(* IEC 61131-3 sources: llm-plc-st-eval/codesys/dobles/I8, 8 files *)

(* ---- 01_Correcta.st ---- *)
(* DOBLE DE PRUEBA I8/Correcta - NO ES CORPUS. Esperado: veredicto 1 *)
FUNCTION_BLOCK FB_Compresor
VAR_INPUT
    pOilOk : BOOL;
    tempOk : BOOL;
    sinAlm : BOOL;
    btnMarcha : BOOL;
    btnParo : BOOL;
END_VAR
VAR_OUTPUT
    comp : BOOL;
    causaBloqueo : INT;
END_VAR
VAR
    tOil : TON;
    fMarcha : R_TRIG;
    oil : BOOL;
    perm : BOOL;
    lat : BOOL;
    pet : BOOL;
END_VAR
tOil(IN := pOilOk, PT := T#3S);
oil := tOil.Q;
IF NOT oil THEN
    causaBloqueo := 1;
ELSIF NOT tempOk THEN
    causaBloqueo := 2;
ELSIF NOT sinAlm THEN
    causaBloqueo := 3;
ELSE
    causaBloqueo := 0;
END_IF
perm := causaBloqueo = 0;
fMarcha(CLK := btnMarcha);
IF btnParo OR NOT perm THEN
    comp := FALSE;
ELSIF fMarcha.Q THEN
    comp := TRUE;
END_IF
END_FUNCTION_BLOCK

(* ---- 02_SinTemporizacionAceite.st ---- *)
(* DOBLE DE PRUEBA I8/SinTemporizacionAceite - NO ES CORPUS. Esperado: veredicto 2, falla en el paso 1 *)
FUNCTION_BLOCK FB_Compresor
VAR_INPUT
    pOilOk : BOOL;
    tempOk : BOOL;
    sinAlm : BOOL;
    btnMarcha : BOOL;
    btnParo : BOOL;
END_VAR
VAR_OUTPUT
    comp : BOOL;
    causaBloqueo : INT;
END_VAR
VAR
    tOil : TON;
    fMarcha : R_TRIG;
    oil : BOOL;
    perm : BOOL;
    lat : BOOL;
    pet : BOOL;
END_VAR
oil := pOilOk;
IF NOT oil THEN
    causaBloqueo := 1;
ELSIF NOT tempOk THEN
    causaBloqueo := 2;
ELSIF NOT sinAlm THEN
    causaBloqueo := 3;
ELSE
    causaBloqueo := 0;
END_IF
perm := causaBloqueo = 0;
fMarcha(CLK := btnMarcha);
IF btnParo OR NOT perm THEN
    comp := FALSE;
ELSIF fMarcha.Q THEN
    comp := TRUE;
END_IF
END_FUNCTION_BLOCK

(* ---- 03_RearranqueAutomatico.st ---- *)
(* DOBLE DE PRUEBA I8/RearranqueAutomatico - NO ES CORPUS. Esperado: veredicto 2, falla en el paso 6 *)
FUNCTION_BLOCK FB_Compresor
VAR_INPUT
    pOilOk : BOOL;
    tempOk : BOOL;
    sinAlm : BOOL;
    btnMarcha : BOOL;
    btnParo : BOOL;
END_VAR
VAR_OUTPUT
    comp : BOOL;
    causaBloqueo : INT;
END_VAR
VAR
    tOil : TON;
    fMarcha : R_TRIG;
    oil : BOOL;
    perm : BOOL;
    lat : BOOL;
    pet : BOOL;
END_VAR
tOil(IN := pOilOk, PT := T#3S);
oil := tOil.Q;
IF NOT oil THEN
    causaBloqueo := 1;
ELSIF NOT tempOk THEN
    causaBloqueo := 2;
ELSIF NOT sinAlm THEN
    causaBloqueo := 3;
ELSE
    causaBloqueo := 0;
END_IF
perm := causaBloqueo = 0;
fMarcha(CLK := btnMarcha);
lat := (lat OR fMarcha.Q) AND NOT btnParo;
comp := lat AND perm;
END_FUNCTION_BLOCK

(* ---- 04_MarchaPrioritaria.st ---- *)
(* DOBLE DE PRUEBA I8/MarchaPrioritaria - NO ES CORPUS. Esperado: veredicto 2, falla en el paso 7 *)
FUNCTION_BLOCK FB_Compresor
VAR_INPUT
    pOilOk : BOOL;
    tempOk : BOOL;
    sinAlm : BOOL;
    btnMarcha : BOOL;
    btnParo : BOOL;
END_VAR
VAR_OUTPUT
    comp : BOOL;
    causaBloqueo : INT;
END_VAR
VAR
    tOil : TON;
    fMarcha : R_TRIG;
    oil : BOOL;
    perm : BOOL;
    lat : BOOL;
    pet : BOOL;
END_VAR
tOil(IN := pOilOk, PT := T#3S);
oil := tOil.Q;
IF NOT oil THEN
    causaBloqueo := 1;
ELSIF NOT tempOk THEN
    causaBloqueo := 2;
ELSIF NOT sinAlm THEN
    causaBloqueo := 3;
ELSE
    causaBloqueo := 0;
END_IF
perm := causaBloqueo = 0;
fMarcha(CLK := btnMarcha);
IF fMarcha.Q AND perm THEN
    comp := TRUE;
ELSIF btnParo OR NOT perm THEN
    comp := FALSE;
END_IF
END_FUNCTION_BLOCK

(* ---- 05_ArrancaPorNivel.st ---- *)
(* DOBLE DE PRUEBA I8/ArrancaPorNivel - NO ES CORPUS. Esperado: veredicto 2, falla en el paso 8 *)
FUNCTION_BLOCK FB_Compresor
VAR_INPUT
    pOilOk : BOOL;
    tempOk : BOOL;
    sinAlm : BOOL;
    btnMarcha : BOOL;
    btnParo : BOOL;
END_VAR
VAR_OUTPUT
    comp : BOOL;
    causaBloqueo : INT;
END_VAR
VAR
    tOil : TON;
    fMarcha : R_TRIG;
    oil : BOOL;
    perm : BOOL;
    lat : BOOL;
    pet : BOOL;
END_VAR
tOil(IN := pOilOk, PT := T#3S);
oil := tOil.Q;
IF NOT oil THEN
    causaBloqueo := 1;
ELSIF NOT tempOk THEN
    causaBloqueo := 2;
ELSIF NOT sinAlm THEN
    causaBloqueo := 3;
ELSE
    causaBloqueo := 0;
END_IF
perm := causaBloqueo = 0;
fMarcha(CLK := btnMarcha);
comp := (comp OR btnMarcha) AND perm AND NOT btnParo;
END_FUNCTION_BLOCK

(* ---- 06_CausaPrioridadInvertida.st ---- *)
(* DOBLE DE PRUEBA I8/CausaPrioridadInvertida - NO ES CORPUS. Esperado: veredicto 2, falla en el paso 0 *)
FUNCTION_BLOCK FB_Compresor
VAR_INPUT
    pOilOk : BOOL;
    tempOk : BOOL;
    sinAlm : BOOL;
    btnMarcha : BOOL;
    btnParo : BOOL;
END_VAR
VAR_OUTPUT
    comp : BOOL;
    causaBloqueo : INT;
END_VAR
VAR
    tOil : TON;
    fMarcha : R_TRIG;
    oil : BOOL;
    perm : BOOL;
    lat : BOOL;
    pet : BOOL;
END_VAR
tOil(IN := pOilOk, PT := T#3S);
oil := tOil.Q;
IF NOT sinAlm THEN
    causaBloqueo := 3;
ELSIF NOT tempOk THEN
    causaBloqueo := 2;
ELSIF NOT oil THEN
    causaBloqueo := 1;
ELSE
    causaBloqueo := 0;
END_IF
perm := causaBloqueo = 0;
fMarcha(CLK := btnMarcha);
IF btnParo OR NOT perm THEN
    comp := FALSE;
ELSIF fMarcha.Q THEN
    comp := TRUE;
END_IF
END_FUNCTION_BLOCK

(* ---- 07_AceiteNoContinuo.st ---- *)
(* DOBLE DE PRUEBA I8/AceiteNoContinuo - NO ES CORPUS. Esperado: veredicto 2, falla en el paso 12 *)
FUNCTION_BLOCK FB_Compresor
VAR_INPUT
    pOilOk : BOOL;
    tempOk : BOOL;
    sinAlm : BOOL;
    btnMarcha : BOOL;
    btnParo : BOOL;
END_VAR
VAR_OUTPUT
    comp : BOOL;
    causaBloqueo : INT;
END_VAR
VAR
    tOil : TON;
    fMarcha : R_TRIG;
    oil : BOOL;
    perm : BOOL;
    lat : BOOL;
    pet : BOOL;
END_VAR
tOil(IN := pOilOk, PT := T#3S);
oil := oil OR tOil.Q;
IF NOT oil THEN
    causaBloqueo := 1;
ELSIF NOT tempOk THEN
    causaBloqueo := 2;
ELSIF NOT sinAlm THEN
    causaBloqueo := 3;
ELSE
    causaBloqueo := 0;
END_IF
perm := causaBloqueo = 0;
fMarcha(CLK := btnMarcha);
IF btnParo OR NOT perm THEN
    comp := FALSE;
ELSIF fMarcha.Q THEN
    comp := TRUE;
END_IF
END_FUNCTION_BLOCK

(* ---- 08_PeticionMemorizada.st ---- *)
(* DOBLE DE PRUEBA I8/PeticionMemorizada - NO ES CORPUS. Esperado: veredicto 2, falla en el paso 14 *)
FUNCTION_BLOCK FB_Compresor
VAR_INPUT
    pOilOk : BOOL;
    tempOk : BOOL;
    sinAlm : BOOL;
    btnMarcha : BOOL;
    btnParo : BOOL;
END_VAR
VAR_OUTPUT
    comp : BOOL;
    causaBloqueo : INT;
END_VAR
VAR
    tOil : TON;
    fMarcha : R_TRIG;
    oil : BOOL;
    perm : BOOL;
    lat : BOOL;
    pet : BOOL;
END_VAR
tOil(IN := pOilOk, PT := T#3S);
oil := tOil.Q;
IF NOT oil THEN
    causaBloqueo := 1;
ELSIF NOT tempOk THEN
    causaBloqueo := 2;
ELSIF NOT sinAlm THEN
    causaBloqueo := 3;
ELSE
    causaBloqueo := 0;
END_IF
perm := causaBloqueo = 0;
fMarcha(CLK := btnMarcha);
pet := (pet OR fMarcha.Q) AND NOT btnParo;
IF btnParo OR (comp AND NOT perm) THEN
    comp := FALSE;
    pet := FALSE;
ELSIF pet AND perm THEN
    comp := TRUE;
END_IF
END_FUNCTION_BLOCK
